// TIA Portal V17 export
// export: Created 2026-11-08T05:50:29.1346515Z, ExportSetting WithDefaults, DisplayName Totally Integrated Automation Portal, DisplayVersion V17, DisplayName TIA Portal Openness, DisplayVersion V17, DisplayName TIA Portal Version Control Interface, DisplayVersion V17, DisplayName STEP 7 Professional, DisplayVersion V17, DisplayName STEP 7 Safety, DisplayVersion V17, DisplayName WinCC Professional, DisplayVersion V17
FUNCTION_BLOCK "FB_Mando_Motor"   // FB1, LAD
TITLE = Mando del motor: pulsadores + HMI
{ S7_Optimized_Access := 'TRUE' }
VERSION : 0.1
// Une pulsadores físicos y botones HMI. Reset = botón RESET de la HMI o mantener MARCHA 3 s.
// stored: AutoNumber true, IsIECCheckEnabled false, IsRetainMemResEnabled false, MemoryReserve 100, SetENOAutomatically false, UDAEnableTagReadback false
   VAR_INPUT
      PB_Marcha : Bool;   // Pulsador MARCHA (NA)
      PB_Paro : Bool;   // Pulsador PARO: 1 = pulsado
      Termico_Falla : Bool;   // Relé térmico: 1 = disparado
      HMI_Marcha : Bool;
      HMI_Paro : Bool;
      HMI_Reset : Bool;
   END_VAR
   VAR_OUTPUT
      Marcha : Bool;
      Paro : Bool;
      Termico_OK : Bool;
      Reset : Bool;
   END_VAR
   VAR
      T_Reset : TON_TIME;   // Tiempo de MARCHA mantenida
      Reset_Mantenido : Bool;   // MARCHA mantenida 3 s
   END_VAR
BEGIN

REGION Network 1: Marcha
   // Pulsador físico o botón de la HMI.
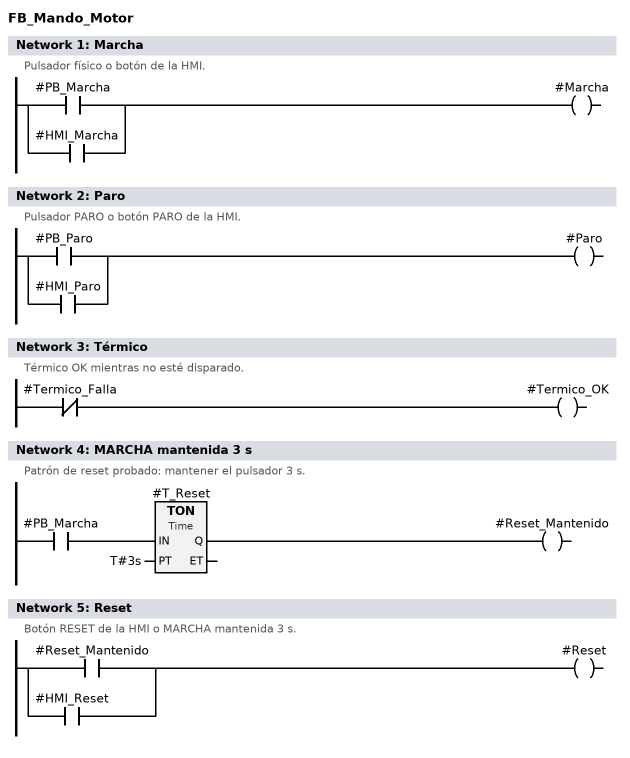
   RUNG wire#powerrail
      Contact( #PB_Marcha )
      wire#w1
      Coil( #Marcha )
   END_RUNG
   RUNG wire#powerrail
      Contact( #HMI_Marcha )
   END_RUNG wire#w1
   // the same network as SCL:
   #Marcha := #PB_Marcha OR #HMI_Marcha;
END_REGION

REGION Network 2: Paro
   // Pulsador PARO o botón PARO de la HMI.
   RUNG wire#powerrail
      Contact( #PB_Paro )
      wire#w1
      Coil( #Paro )
   END_RUNG
   RUNG wire#powerrail
      Contact( #HMI_Paro )
   END_RUNG wire#w1
   // the same network as SCL:
   #Paro := #PB_Paro OR #HMI_Paro;
END_REGION

REGION Network 3: Térmico
   // Térmico OK mientras no esté disparado.
   RUNG wire#powerrail
      I_Contact( #Termico_Falla )
      Coil( #Termico_OK )
   END_RUNG
   // the same network as SCL:
   #Termico_OK := NOT #Termico_Falla;
END_REGION

REGION Network 4: MARCHA mantenida 3 s
   // Patrón de reset probado: mantener el pulsador 3 s.
   RUNG wire#powerrail
      Contact( #PB_Marcha )
      { S7_Templates := "time_type := Time" } #T_Reset.TON(pt := T#3s, et =>)
      Coil( #Reset_Mantenido )
   END_RUNG
   // the same network as SCL:
   #T_Reset(IN := #PB_Marcha, PT := T#3s);   // TON
   #Reset_Mantenido := #T_Reset.Q;
END_REGION

REGION Network 5: Reset
   // Botón RESET de la HMI o MARCHA mantenida 3 s.
   RUNG wire#powerrail
      Contact( #Reset_Mantenido )
      wire#w1
      Coil( #Reset )
   END_RUNG
   RUNG wire#powerrail
      Contact( #HMI_Reset )
   END_RUNG wire#w1
   // the same network as SCL:
   #Reset := #Reset_Mantenido OR #HMI_Reset;
END_REGION
END_FUNCTION_BLOCK
